Fanuc KAREL source: KT00105.KL

PROGRAM KT00105
%NOLOCKGROUP
VAR
  R1: REAL
  I2: INTEGER
  OUT: INTEGER
BEGIN
  R1 = 2.0
    I2 = 3
  OUT = R1 / I2
END KT00105
